TYPE ST_TouchProbeRenishawStatus :
STRUCT
	bProbeStatus1					:BOOL;			(* Probe status 1 *)
	bLowBattery						:BOOL;			(* Low battery  *)
	bError							:BOOL;			(* Error  *)
END_STRUCT
END_TYPE

(* stored: Version 1.1.0.1, ProductVersion 3.1.4024.15
   DUT ST_TouchProbeRenishawStatus: Id {1e71fcd9-3937-453b-a835-93c4283a5fcc} *)
